FUNCTION_BLOCK FB_MoveToNearestClosed
VAR_OUTPUT
    Closed   : BOOL;
END_VAR
VAR
    iMotionStage 		: I_MotionStage;
    fEndpointPositive  : LREAL :=  11.25;
    fEndpointNegative  : LREAL := -11.25;
    fTarget            : LREAL := 0.0;
    bStarted: BOOL;
END_VAR

Closed := FALSE;
IF 	bStarted THEN
    IF iMotionStage.MotionStatus.bDone THEN
        Closed := TRUE;
        bStarted := FALSE;
    END_IF
END_IF

//FB_Init is always available implicitly and it is used primarily for initialization.
//The return value is not evaluated. For a specific influence, you can also declare the
//methods explicitly and provide additional code there with the standard initialization
//code. You can evaluate the return value.
METHOD FB_Init: BOOL
VAR_INPUT
    bInitRetains: BOOL; // TRUE: the retain variables are initialized (reset warm / reset cold)
    bInCopyCode: BOOL;  // TRUE: the instance will be copied to the copy code afterward (online change)
    iMotionStage : I_MotionStage;
END_VAR
THIS^.iMotionStage := iMotionStage ;
END_METHOD

METHOD Start
// Choose closest endpoint
IF ABS(iMotionStage.MotionStatus.fActPosition - fEndpointPositive) < ABS(iMotionStage.MotionStatus.fActPosition - fEndpointNegative) THEN
    fTarget := fEndpointPositive;
ELSE
    fTarget := fEndpointNegative;
END_IF
// Issue move command
iMotionStage.AbsoluteMove(
   Position     := fTarget,
   Velocity     := iMotionStage.MotionCmd.fVelocity,
   Acceleration := iMotionStage.MotionCmd.fAcceleration,
   Deceleration := iMotionStage.MotionCmd.fDeceleration
);

bStarted := TRUE;
END_METHOD

END_FUNCTION_BLOCK

(* stored: Version 1.1.0.1
   POU FB_MoveToNearestClosed: Id {6ed107c2-bebb-4576-9274-e415e2ee6172}, SpecialFunc None
   Method FB_Init: Id {d19b4830-b739-4f72-bb4a-99a9c85524b7}
   Method Start: Id {70fa49d8-d54b-4879-afbc-54860b8a35fc} *)
